Universal Robots PolyScope program: TgtProg.urp

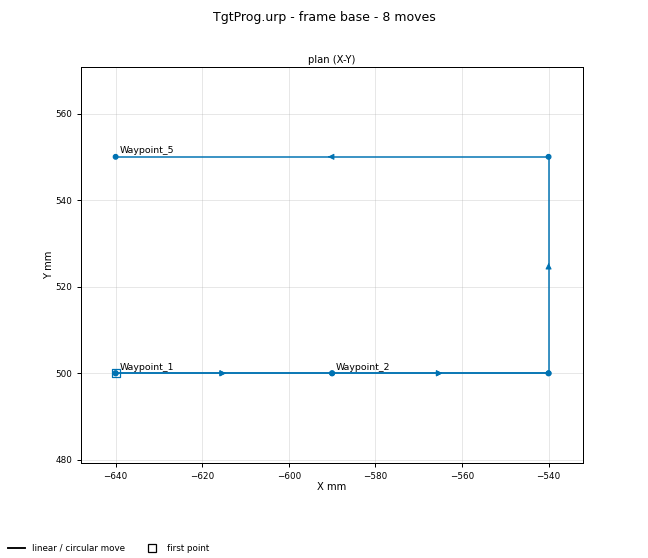
[picture p0: tool path of TgtProg.urp in frame base, 8 of 9 moves have a stored position in this frame; points joined in program order, loops and branches not executed]
Program TgtProg (createdIn=3.0.0 lastSavedIn=3.0.0 directory=/programs installation=default)
Robot Program (runOnlyOnce=true motionType=MoveJ speed=1.047198 acceleration=1.396263 useActiveTCP=false)
  'Program generated by RoboDK v6.0.7 for UR10 on XX/XX/XXXX 18:00:00'
  'Using nominal kinematics.'
  'Using TCP T: p[0.000000, 0.000000, 0.100000, 0.000000, 0.000000, 0.000000]'
  Script: set_tcp(p[0.000000, 0.000000, 0.100000, 0.000000, 0.000000, 0.000000])
  MoveL speed 250 mm/s, acceleration 1200 mm/s^2 (useActiveTCP=true)
    Waypoint Waypoint_1: TCP in base x=-640 y=500 z=370 mm, rx=0.732 ry=2.1859 rz=-0.5703 rad; joints [0, -10, 20, 0, 30, 0] deg; flange x=-691.14 y=559.411 z=432.089 mm, rx=0.732 ry=2.1859 rz=-0.5703 rad
  MoveL speed 100 mm/s, acceleration 1200 mm/s^2 (useActiveTCP=true)
    Waypoint Waypoint_2: TCP in base x=-590 y=500 z=370 mm, rx=0.732 ry=2.1859 rz=-0.5703 rad; joints [0, -10, 20, 0, 30, 0] deg; flange x=-641.14 y=559.411 z=432.089 mm, rx=0.732 ry=2.1859 rz=-0.5703 rad
  MoveL speed 100 mm/s, acceleration 1200 mm/s^2 (useActiveTCP=true)
    Waypoint Waypoint_3: TCP in base x=-540 y=500 z=370 mm, rx=0.732 ry=2.1859 rz=-0.5703 rad; joints [0, -10, 20, 0, 30, 0] deg; flange x=-591.14 y=559.411 z=432.089 mm, rx=0.732 ry=2.1859 rz=-0.5703 rad
    Waypoint Waypoint_4: motionParameters(blendRadius=0 jointSpeed=0.75 jointAcceleration=1.2 cartesianSpeed=0.1 cartesianAcceleration=0.5); TCP in base x=-540 y=550 z=370 mm, rx=0.732 ry=2.1859 rz=-0.5703 rad; joints [0, -10, 20, 0, 30, 0] deg; flange x=-591.14 y=609.411 z=432.089 mm, rx=0.732 ry=2.1859 rz=-0.5703 rad
  'note'
  MoveL speed 100 mm/s, acceleration 500 mm/s^2 (useActiveTCP=true)
    Waypoint Waypoint_5: TCP in base x=-640 y=550 z=370 mm, rx=0.732 ry=2.1859 rz=-0.5703 rad; joints [0, -10, 20, 0, 30, 0] deg; flange x=-691.14 y=609.411 z=432.089 mm, rx=0.732 ry=2.1859 rz=-0.5703 rad
    Waypoint Waypoint_6: position(joints=0.174533, -0.174533, 0.349066, 0.000000, 0.523599, 0.087266)
    Waypoint Waypoint_7: TCP in base x=-640 y=500 z=370 mm, rx=0.732 ry=2.1859 rz=-0.5703 rad; joints [0, -10, 20, 0, 30, 0] deg; flange x=-691.14 y=559.411 z=432.089 mm, rx=0.732 ry=2.1859 rz=-0.5703 rad
    Waypoint Waypoint_8: motionParameters(blendRadius=0.002); TCP in base x=-590 y=500 z=370 mm, rx=0.732 ry=2.1859 rz=-0.5703 rad; joints [0, -10, 20, 0, 30, 0] deg; flange x=-641.14 y=559.411 z=432.089 mm, rx=0.732 ry=2.1859 rz=-0.5703 rad
    Waypoint Waypoint_9: motionParameters(blendRadius=0.002 jointSpeed=0.349066 jointAcceleration=1.2 cartesianSpeed=0.1 cartesianAcceleration=0.5); TCP in base x=-540 y=500 z=370 mm, rx=0.732 ry=2.1859 rz=-0.5703 rad; joints [0, -10, 20, 0, 30, 0] deg; flange x=-591.14 y=559.411 z=432.089 mm, rx=0.732 ry=2.1859 rz=-0.5703 rad
